// TIA Portal V21 export
Screen "T11_LampAlarm"  1024x768, Number=31
  ScreenLayer 
    Rectangle "P_LampAlarm" at 0,0 size 100x30
      AppearanceAnimation   AnimationMode=Range, Tag=LampAlarm
        AppearanceAnimationRange 
        AppearanceAnimationRange   Range=1
